(* IEC 61131-3 sources: STEPROBOT/docs/welder_r6_4/plc, 4 files *)

(* ---- GVL_WelderBridge.st ---- *)
{attribute 'qualified_only'}
VAR_GLOBAL PERSISTENT RETAIN
    // AC802 fixed MW registers require both persistence attributes.
    aCommand AT %MW7000 : ARRAY[0..31] OF WORD;
    wHeartbeat AT %MW7064 : WORD;
    aStatus AT %MW7200 : ARRAY[0..63] OF WORD;
END_VAR

VAR_GLOBAL
    // Local commissioning inputs; never write these over the PC command channel.
    xMappingConfirmed : BOOL := FALSE;
    xWeldPermit : BOOL := FALSE;
    // Drive from the real EtherCAT slave OP / working-counter-valid signal.
    // A constant TRUE is not a valid connection-health signal.
    xPdoOperational : BOOL := FALSE;
END_VAR

(* ---- GVL_Welders.st ---- *)
(* Reused legacy EtherCAT PDO variables. No fixed addresses or retained process outputs.
   Old Dxxx comments describe the source only; PC uses HR7000 / HR7200. *)
VAR_GLOBAL
    (* EtherCAT输出 → 焊机输入数据区 (32字节) *)
    g_byWeldOut : ARRAY[0..31] OF BYTE;
    (* EtherCAT输入 ← 焊机输出数据区 (32字节) *)
    g_byWeldIn : ARRAY[0..31] OF BYTE;

    (*
     * EtherCAT 映射别名。
     * InoProShop 的 I/O 映射器要求变量是单一标识符，不接受数组下标；
     * CommPoll 在这些别名与协议数组之间逐周期同步，协议字节编号保持不变。
     *)
    g_byWeldOutMap01 : BYTE;
    g_byWeldOutMap02 : BYTE;
    g_byWeldOutMap03 : BYTE;
    g_byWeldOutMap04 : BYTE;
    g_byWeldOutMap05 : BYTE;
    g_byWeldOutMap06 : BYTE;
    g_byWeldOutMap07 : BYTE;
    g_byWeldOutMap08 : BYTE;
    g_byWeldOutMap09 : BYTE;
    g_byWeldOutMap10 : BYTE;
    g_byWeldOutMap11 : BYTE;
    g_byWeldOutMap12 : BYTE;
    g_byWeldOutMap13 : BYTE;
    g_byWeldOutMap14 : BYTE;
    g_byWeldOutMap15 : BYTE;
    g_byWeldOutMap16 : BYTE;
    g_byWeldOutMap17 : BYTE;
    g_byWeldOutMap18 : BYTE;
    g_byWeldOutMap19 : BYTE;
    g_byWeldOutMap20 : BYTE;
    g_byWeldOutMap21 : BYTE;
    g_byWeldOutMap22 : BYTE;
    g_byWeldOutMap23 : BYTE;
    g_byWeldOutMap24 : BYTE;
    g_byWeldOutMap25 : BYTE;
    g_byWeldOutMap26 : BYTE;
    g_byWeldOutMap27 : BYTE;
    g_byWeldOutMap28 : BYTE;
    g_byWeldOutMap29 : BYTE;
    g_byWeldOutMap30 : BYTE;
    g_byWeldOutMap31 : BYTE;
    g_byWeldOutMap32 : BYTE;

    g_byWeldInMap01 : BYTE;
    g_byWeldInMap02 : BYTE;
    g_byWeldInMap03 : BYTE;
    g_byWeldInMap04 : BYTE;
    g_byWeldInMap05 : BYTE;
    g_byWeldInMap06 : BYTE;
    g_byWeldInMap07 : BYTE;
    g_byWeldInMap08 : BYTE;
    g_byWeldInMap09 : BYTE;
    g_byWeldInMap10 : BYTE;
    g_byWeldInMap11 : BYTE;
    g_byWeldInMap12 : BYTE;
    g_byWeldInMap13 : BYTE;
    g_byWeldInMap14 : BYTE;
    g_byWeldInMap15 : BYTE;
    g_byWeldInMap16 : BYTE;
    g_byWeldInMap17 : BYTE;
    g_byWeldInMap18 : BYTE;
    g_byWeldInMap19 : BYTE;
    g_byWeldInMap20 : BYTE;
    g_byWeldInMap21 : BYTE;
    g_byWeldInMap22 : BYTE;
    g_byWeldInMap23 : BYTE;
    g_byWeldInMap24 : BYTE;
    g_byWeldInMap25 : BYTE;
    g_byWeldInMap26 : BYTE;
    g_byWeldInMap27 : BYTE;
    g_byWeldInMap28 : BYTE;
    g_byWeldInMap29 : BYTE;
    g_byWeldInMap30 : BYTE;
    g_byWeldInMap31 : BYTE;
    g_byWeldInMap32 : BYTE;

	(* D520 | 激光距离 (原始INT值, 从%IW50读取) *)
	(* --- 激光距离原始值 --- *)
	g_iLaserDistanceRaw : INT;
END_VAR

VAR_GLOBAL

(* D300 | 控制标志位打包字 (PC通过Modbus读写, CommPoll每周期双向映射) *)
g_wWeldCtrlWord : UINT := 0;

(* D300 bit0 | 独立BOOL | 开始焊接 1=起弧 0=停弧 [危险, 高有效] *)
g_wWeldOn : BOOL := FALSE;

(* D300 bit1 | 独立BOOL | 机器人准备好, 高有效 *)
g_wRobotReady : BOOL := FALSE;
(* D300 bit2 | 独立BOOL | 检气, 高有效 *)
g_wGasCheck : BOOL := FALSE;

(* D300 bit3 | 独立BOOL | 热丝电源使能 1=ON 0=OFF *)
g_bHotWireEnable : BOOL := FALSE;

(* D300 bit4 | 独立BOOL | 热丝工作模式 0=DC 1=AC *)
g_bHotWireACMode : BOOL := FALSE;

(* D300 bit7 | 独立BOOL | 高频有无 0=高频 1=提升 *)
g_bHighFreqDisable : BOOL := FALSE;

(* D300 bit8 | 独立BOOL | 焊枪模式 0=水冷 1=气冷 *)
g_bGunCoolMode : BOOL := FALSE;

(* D302 | 协议Byte0 bit3-4 | 焊机操作模式 0=两步 1=四步 2=反复 *)
g_wWeldOperMode : UINT := 0;

(* D304 | 协议Byte0 bit5-7 | 焊机工作模式 0=直流恒流 1=直流脉冲 2=交流恒流 *)
(*                           3=交流脉冲 4=直流手弧焊 *)
g_wWeldWorkMode : UINT := 1;

(* D306 | 协议Byte11 | 通讯异常标志, 控制器填充, 默认0 *)
g_wCommErrorFlag : BYTE;

(* D414 | 协议Byte2 bit0-7 | 热丝频率, 范围20~100, 对应20~100Hz (直通) *)
g_wHotWireFreq : UINT := 50;

(* D416 | 协议Byte3 bit0-7 | 热丝电流给定, 范围0~200, 对应0~200A (直通) *)
g_wHotWireCurrent : UINT := 150;

(* D400 | 协议Byte4-5 | 给定电流, 实际A, 例: 100.0表示100.0A *)
(* CommPoll内部 ×10 → 协议值(范围40~4000, 对应4.0~400.0A), 占D400-D401 *)
g_wWeldCurrent : REAL := 100.0;

(* Local wire-feed axis parameters. Speeds are mm/s; delays are seconds.
   D412 and D1202 set the same automatic speed; a changed D1202 has priority.
   D410 > 0 overrides D2104 for axis 4 jog; zero uses D2104 for compatibility. *)
g_rWireStartDelay : REAL := 0.0;
g_rWireStopDelay : REAL := 0.0;
g_rWireJogSpeed : REAL := 0.0;
g_rWireAutoSpeed : REAL := 0.0;

(* D420 | 协议Byte13-14 | 前气时间, 实际s, 例: 5.0表示5.00s *)
(* CommPoll内部 ×100 → 协议值(范围1~999, 对应0.01~9.99s), 占D420-D421 *)
g_wFrontGasTime : REAL := 0.01;

(* D422 | 协议Byte15-16 | 延气时间, 实际s, 例: 3.0表示3.0s *)
(* CommPoll内部 ×10 → 协议值(范围1~600, 对应0.1~60.0s), 占D422-D423 *)
g_wTailGasTime : REAL := 0.2;

(* D424 | 协议Byte17 bit0-7 | 爬升时间, 实际s, 例: 5.0表示5.0s *)
(* CommPoll内部 ×10 → 协议值(范围1~100, 对应0.1~10.0s), 占D424-D425 *)
g_wRampUpTime : REAL := 0.5;

(* D426 | 协议Byte18 bit0-7 | 衰减时间, 实际s, 例: 5.0表示5.0s *)
(* CommPoll内部 ×10 → 协议值(范围1~150, 对应0.1~15.0s) *)
g_wRampDownTime : REAL := 0.2;

(* D428 | 协议Byte19 bit0-7 | 脉冲频率, 实际Hz, 例: 5.0表示5.0Hz *)
(* CommPoll内部 ×10 → 协议值(范围2~200, 对应0.2~20.0Hz), 占D428-D429 *)
g_wPulseFreq : REAL := 0.5;

(* D430 | 协议Byte20+22 bit4-7 | 占空比, 实际百分比, 例: 50.0表示50.0% *)
(* CommPoll内部 ×10 → 协议值(范围1~999, 对应0.1%~99.9%), 占D430-D431 *)
g_wDutyCycle : REAL := 50.0;

(* D432 | 协议Byte21+22 bit0-3 | 峰值电流, 实际A, 例: 150.0表示150.0A *)
(* CommPoll内部 ×10 → 协议值(范围50~4000, 对应5.0~400.0A), 占D432-D433 *)
g_wPeakCurrent : REAL := 100.0;

(* D434 | 协议Byte23-24 | 基值电流, 实际A, 例: 30.0表示30.0A *)
(* CommPoll内部 ×10 → 协议值(范围50~4000, 对应5.0~400.0A), 占D434-D435 *)
g_wBaseCurrent : REAL := 30.0;

(* D436 | 协议Byte25-26 | 起弧电流, 实际A, 例: 100.0表示100.0A *)
(* CommPoll内部 ×10 → 协议值(范围50~4000, 对应5.0~400.0A), 占D436-D437 *)
(* --- 协议 Byte 25-26: 起弧电流 (2字节小端, 低字节在前) --- *)
g_wArcStartCurrent : REAL := 5.0;

(* D438 | 协议Byte27-28 | 收弧电流, 实际A, 例: 100.0表示100.0A *)
(* CommPoll内部 ×10 → 协议值(范围50~4000, 对应5.0~400.0A), 占D438-D439 *)
(* --- 协议 Byte 27-28: 收弧电流 (2字节小端, 低字节在前) --- *)
g_wArcEndCurrent : REAL := 5.0;

(* D440 | 协议Byte29 bit0-7 | 交流频率, 范围40~250, 对应40~250Hz (直通) *)
(* --- 协议 Byte 29: 交流频率 --- *)
g_wACFreq : UINT := 40;

(* D442 | 协议Byte30 bit0-7 | 清理比例, 范围90~180, 对应40~-50 *)
(* 协议转换: Byte30 = -1 × D442 + 130 *)
(* 例: D442=90 → Byte30=40, D442=130 → Byte30=0, D442=180 → Byte30=-50 *)
(* --- 协议 Byte 30: 清理比例 --- *)
g_wCleanRatio : UINT := 90;

(* D444 | 协议Byte31 bit0-7 | 交流偏置, 范围90~180, 对应40~-50 *)
(* 协议转换: Byte31 = -1 × D444 + 130 *)
(* 例: D444=90 → Byte31=40, D444=130 → Byte31=0, D444=180 → Byte31=-50 *)
(* --- 协议 Byte 31: 交流偏置 --- *)
g_wACBias : UINT := 90;

(* D308 | 输入状态打包字 (PC通过Modbus读取, CommPoll每周期从独立BOOL组装) *)
g_wWeldStatusWord : UINT;

(* D308 bit0 | 独立BOOL | 引弧成功, 高有效 *)
g_bWeldArcOK : BOOL;

(* D308 bit1 | 独立BOOL | 焊机准备好, 高有效 *)
g_bWeldReady : BOOL;

(* D308 bit2 | 独立BOOL | 电流有无, 高有效 *)
g_bWeldHasCurrent : BOOL;

(* D308 bit3 | 独立BOOL | 焊枪开关异常, 高有效 *)
g_bGunSwitchFault : BOOL;

(* D308 bit4 | 独立BOOL | 焊机热保护, 高有效 *)
g_bWeldThermalProtect : BOOL;

(* D308 bit5 | 独立BOOL | 缺水保护, 高有效 *)
g_bWaterProtect : BOOL;

(* D308 bit6 | 独立BOOL | 热丝电源热保护, 高有效 *)
g_bWirePSThermal : BOOL;

(* D308 bit7 | 独立BOOL | 热丝电源通讯保护, 高有效, 控制器填充 *)
g_bWirePSCommFault : BOOL;

(* D308 bit8 | 独立BOOL | 组合报警, 包含焊枪开关/热保护/缺水/热丝电源故障 *)
g_bWeldFault : BOOL;

(* D500 | 焊机输入状态字 (16位打包, 详见位域定义) *)
g_wWeldInStatus : UINT;

(* D502-D503 | 协议输入Byte4-5 | 实际焊接电压, 0.1V分辨率 *)
(* --- 协议输入 Byte 4-5: 实际焊接电压 (2字节小端, 0.1V分辨率) --- *)
(* 范围: 0~1000 → 0~100.0V *)
g_rWeldVoltageAct : REAL;

(* D506-D507 | 协议输入Byte6-7 | 实际焊接电流, 0.1A分辨率 *)
(* --- 协议输入 Byte 6-7: 实际焊接电流 (2字节小端, 0.1A分辨率) --- *)
(* 范围: 0~400 → 0~400A *)
g_rWeldCurrentAct : REAL;

(* D510-D511 | 协议输入Byte8-9 | 实际热丝焊接电流, 10A分辨率 *)
(* --- 协议输入 Byte 8-9: 实际热丝焊接电流 (2字节小端, 10A分辨率) --- *)
(* 范围: 0~20 → 0~200A *)
g_rHotWireCurrentAct : REAL;

(* D518 | 协议输入Byte1原始值 | 报警码, 报警时记录协议输入Byte1原始值 *)
(* --- 报警原始字节 --- *)
g_rWeldFaultCode : UINT;

(* D522 | 激光距离 (实际距离mm, 原始值/100+50) *)
(* --- 激光距离实际值 --- *)
g_rLaserDistance : REAL := 50.0;

(* ================================================================= *)
(* 协议输入预留字节 (协议保留, 当前未使用)                               *)
(*   协议输入 Byte 2-3: 预留                                          *)
(*   协议输入 Byte 12:  预留                                          *)
(* ================================================================= *)

END_VAR

(* ---- PRG_WelderBridge.st ---- *)
PROGRAM PRG_WelderBridge
VAR
    aFrame : ARRAY[0..31] OF WORD;
    aParam : ARRAY[0..19] OF WORD;
    uiI : UINT;
    wCheck : WORD;
    uiScan : UINT;
    wPreviousHeartbeat : WORD;
    xHeartbeatSeen : BOOL;
    xHeartbeatEdge : BOOL;
    fbWatchdog : TON;
    xHostFresh : BOOL;
    xBasePermit : BOOL;
    xArcPermit : BOOL;
    xParametersValid : BOOL;
    xWasRunning : BOOL;
    xJobEnded : BOOL;
    udiOwner : UDINT;
    udiCurrentOwner : UDINT;
    udiRequest : UDINT;
    udiLastRequest : UDINT;
    udiRequestOwner : UDINT;
    udiRequestBoot : UDINT;
    udiBoot : UDINT;
    wResult : WORD;
    wError : WORD;
    wOperation : WORD;
    wControl : WORD;
    wApplied : WORD;
END_VAR

// Call once per scan, after PRG_RobotBridge. No other task writes the welder PDOs.
udiBoot := GVL_RobotBridgeRetain.udiBootCounter;
udiCurrentOwner := SHL(WORD_TO_UDINT(GVL_RobotBridge.aHostStatus[15]),16) OR WORD_TO_UDINT(GVL_RobotBridge.aHostStatus[16]);
IF udiCurrentOwner <> udiOwner THEN
    udiOwner := udiCurrentOwner; udiLastRequest := 0; wControl := 0;
    xHeartbeatSeen := FALSE; wPreviousHeartbeat := GVL_WelderBridge.wHeartbeat;
END_IF;
xHeartbeatEdge := GVL_WelderBridge.wHeartbeat <> wPreviousHeartbeat;
IF xHeartbeatEdge THEN
    wPreviousHeartbeat := GVL_WelderBridge.wHeartbeat; xHeartbeatSeen := TRUE;
END_IF;
fbWatchdog(IN := NOT xHeartbeatEdge, PT := T#1200ms);
xHostFresh := xHeartbeatSeen AND NOT fbWatchdog.Q AND GVL_RobotBridge.xHostRegistered AND GVL_RobotBridge.xHostAlive AND (udiOwner <> 0);
xBasePermit := xHostFresh AND GVL_WelderBridge.xMappingConfirmed AND GVL_WelderBridge.xWeldPermit AND GVL_WelderBridge.xPdoOperational
    AND GVL_RobotBridge.xRobotLinkOK AND GVL_RobotBridge.xRemotePermit
    AND NOT GVL_RobotBridge.xStopInterlock AND NOT GVL_RobotBridge.xRobotEmergency AND NOT GVL_RobotBridge.xRobotAlarm;
xArcPermit := xBasePermit AND GVL_RobotBridge.xRobotExternalAuto AND NOT GVL_RobotBridge.xRobotPaused;
xJobEnded := xWasRunning AND NOT GVL_RobotBridge.xRobotRunning;
xWasRunning := GVL_RobotBridge.xRobotRunning;
IF NOT xBasePermit THEN wControl := 0; END_IF;
IF NOT xArcPermit OR xJobEnded THEN wControl := wControl AND WORD#16#0006; END_IF;

// Snapshot the whole FC16 frame, then check checksum, identity and monotonic request.
FOR uiI := 0 TO 31 DO aFrame[uiI] := GVL_WelderBridge.aCommand[uiI]; END_FOR;
udiRequest := SHL(WORD_TO_UDINT(aFrame[2]),16) OR WORD_TO_UDINT(aFrame[3]);
udiRequestOwner := SHL(WORD_TO_UDINT(aFrame[4]),16) OR WORD_TO_UDINT(aFrame[5]);
udiRequestBoot := SHL(WORD_TO_UDINT(aFrame[6]),16) OR WORD_TO_UDINT(aFrame[7]);
wCheck := WORD#16#A55A;
FOR uiI := 0 TO 30 DO wCheck := wCheck XOR aFrame[uiI]; END_FOR;
IF (aFrame[0] = WORD#16#5742) AND (aFrame[1] = WORD#1) AND (wCheck = aFrame[31])
    AND (udiRequestOwner = udiOwner) AND (udiOwner <> 0) AND (udiRequestBoot = udiBoot)
    AND (udiRequest > udiLastRequest) THEN
    udiLastRequest := udiRequest; wOperation := aFrame[8]; wResult := 2; wError := 0;
    IF wOperation = WORD#3 THEN
        wControl := 0; wResult := 1;
    ELSIF NOT xBasePermit THEN
        wError := 1;
    ELSIF wOperation = WORD#1 THEN
        IF (aFrame[9] AND WORD#16#FFF0) <> 0 THEN wError := 2;
        ELSIF ((aFrame[9] AND WORD#16#0009) <> 0) AND NOT xArcPermit THEN wError := 3;
        ELSIF ((aFrame[9] AND WORD#16#0009) <> 0) AND (((aFrame[9] AND WORD#2) = 0) OR NOT GVL_Welders.g_bWeldReady OR GVL_Welders.g_bWeldFault) THEN wError := 4;
        ELSIF ((aFrame[9] AND WORD#1) <> 0) AND ((aFrame[9] AND WORD#4) <> 0) THEN wError := 5;
        ELSE wControl := aFrame[9]; wResult := 1;
        END_IF;
    ELSIF wOperation = WORD#2 THEN
        IF wControl <> 0 THEN wError := 6;
        ELSE
            FOR uiI := 0 TO 19 DO aParam[uiI] := aFrame[10+uiI]; END_FOR;
            xParametersValid := TRUE;
            IF (aParam[0] < WORD#0) OR (aParam[0] > WORD#2) THEN xParametersValid := FALSE; END_IF;
            IF (aParam[1] < WORD#0) OR (aParam[1] > WORD#4) THEN xParametersValid := FALSE; END_IF;
            IF (aParam[2] < WORD#40) OR (aParam[2] > WORD#4000) THEN xParametersValid := FALSE; END_IF;
            IF (aParam[3] < WORD#20) OR (aParam[3] > WORD#100) THEN xParametersValid := FALSE; END_IF;
            IF (aParam[4] < WORD#0) OR (aParam[4] > WORD#200) THEN xParametersValid := FALSE; END_IF;
            IF (aParam[5] < WORD#1) OR (aParam[5] > WORD#999) THEN xParametersValid := FALSE; END_IF;
            IF (aParam[6] < WORD#1) OR (aParam[6] > WORD#600) THEN xParametersValid := FALSE; END_IF;
            IF (aParam[7] < WORD#1) OR (aParam[7] > WORD#100) THEN xParametersValid := FALSE; END_IF;
            IF (aParam[8] < WORD#1) OR (aParam[8] > WORD#150) THEN xParametersValid := FALSE; END_IF;
            IF (aParam[9] < WORD#2) OR (aParam[9] > WORD#200) THEN xParametersValid := FALSE; END_IF;
            IF (aParam[10] < WORD#1) OR (aParam[10] > WORD#999) THEN xParametersValid := FALSE; END_IF;
            IF (aParam[11] < WORD#50) OR (aParam[11] > WORD#4000) THEN xParametersValid := FALSE; END_IF;
            IF (aParam[12] < WORD#50) OR (aParam[12] > WORD#4000) THEN xParametersValid := FALSE; END_IF;
            IF (aParam[13] < WORD#50) OR (aParam[13] > WORD#4000) THEN xParametersValid := FALSE; END_IF;
            IF (aParam[14] < WORD#50) OR (aParam[14] > WORD#4000) THEN xParametersValid := FALSE; END_IF;
            IF (aParam[15] < WORD#40) OR (aParam[15] > WORD#250) THEN xParametersValid := FALSE; END_IF;
            IF (aParam[16] < WORD#90) OR (aParam[16] > WORD#180) THEN xParametersValid := FALSE; END_IF;
            IF (aParam[17] < WORD#90) OR (aParam[17] > WORD#180) THEN xParametersValid := FALSE; END_IF;
            IF (aParam[18] > WORD#7) OR (aParam[19] <> 0) THEN xParametersValid := FALSE; END_IF;
            IF NOT xParametersValid THEN wError := 7;
            ELSE
                GVL_Welders.g_wWeldOperMode := WORD_TO_UINT(aParam[0]);
                GVL_Welders.g_wWeldWorkMode := WORD_TO_UINT(aParam[1]);
                GVL_Welders.g_wWeldCurrent := UINT_TO_REAL(WORD_TO_UINT(aParam[2])) / 10.0;
                GVL_Welders.g_wHotWireFreq := WORD_TO_UINT(aParam[3]);
                GVL_Welders.g_wHotWireCurrent := WORD_TO_UINT(aParam[4]);
                GVL_Welders.g_wFrontGasTime := UINT_TO_REAL(WORD_TO_UINT(aParam[5])) / 100.0;
                GVL_Welders.g_wTailGasTime := UINT_TO_REAL(WORD_TO_UINT(aParam[6])) / 10.0;
                GVL_Welders.g_wRampUpTime := UINT_TO_REAL(WORD_TO_UINT(aParam[7])) / 10.0;
                GVL_Welders.g_wRampDownTime := UINT_TO_REAL(WORD_TO_UINT(aParam[8])) / 10.0;
                GVL_Welders.g_wPulseFreq := UINT_TO_REAL(WORD_TO_UINT(aParam[9])) / 10.0;
                GVL_Welders.g_wDutyCycle := UINT_TO_REAL(WORD_TO_UINT(aParam[10])) / 10.0;
                GVL_Welders.g_wPeakCurrent := UINT_TO_REAL(WORD_TO_UINT(aParam[11])) / 10.0;
                GVL_Welders.g_wBaseCurrent := UINT_TO_REAL(WORD_TO_UINT(aParam[12])) / 10.0;
                GVL_Welders.g_wArcStartCurrent := UINT_TO_REAL(WORD_TO_UINT(aParam[13])) / 10.0;
                GVL_Welders.g_wArcEndCurrent := UINT_TO_REAL(WORD_TO_UINT(aParam[14])) / 10.0;
                GVL_Welders.g_wACFreq := WORD_TO_UINT(aParam[15]);
                GVL_Welders.g_wCleanRatio := WORD_TO_UINT(aParam[16]);
                GVL_Welders.g_wACBias := WORD_TO_UINT(aParam[17]);
                GVL_Welders.g_bHotWireACMode := (aParam[18] AND WORD#1) <> 0;
                GVL_Welders.g_bHighFreqDisable := (aParam[18] AND WORD#2) <> 0;
                GVL_Welders.g_bGunCoolMode := (aParam[18] AND WORD#4) <> 0;
                wResult := 1;
            END_IF;
        END_IF;
    ELSE wError := 8;
    END_IF;
END_IF;
GVL_Welders.g_wWeldOn := (wControl AND WORD#1) <> 0;
GVL_Welders.g_wRobotReady := (wControl AND WORD#2) <> 0;
GVL_Welders.g_wGasCheck := (wControl AND WORD#4) <> 0;
GVL_Welders.g_bHotWireEnable := (wControl AND WORD#8) <> 0;
PRG_WelderIo();
// Same-scan PDO input interlock; never restore an arc after a fault clears.
IF NOT GVL_Welders.g_bWeldReady OR GVL_Welders.g_bWeldFault THEN
    wControl := wControl AND WORD#16#0006;
    GVL_Welders.g_wWeldOn := FALSE; GVL_Welders.g_bHotWireEnable := FALSE;
    GVL_Welders.g_byWeldOutMap01 := GVL_Welders.g_byWeldOutMap01 AND BYTE#16#FE;
    GVL_Welders.g_byWeldOutMap02 := GVL_Welders.g_byWeldOutMap02 AND BYTE#16#FE;
END_IF;
wApplied := wControl;
GVL_Welders.g_wWeldCtrlWord := WORD_TO_UINT(wApplied);
uiScan := uiScan + UINT#1;
GVL_WelderBridge.aStatus[0] := WORD#16#5742;
GVL_WelderBridge.aStatus[1] := 1;
GVL_WelderBridge.aStatus[2] := UINT_TO_WORD(uiScan);
GVL_WelderBridge.aStatus[3] := 1;
IF GVL_WelderBridge.xMappingConfirmed THEN GVL_WelderBridge.aStatus[3] := GVL_WelderBridge.aStatus[3] OR WORD#2; END_IF;
IF GVL_WelderBridge.xPdoOperational THEN GVL_WelderBridge.aStatus[3] := GVL_WelderBridge.aStatus[3] OR WORD#4; END_IF;
IF xBasePermit THEN GVL_WelderBridge.aStatus[3] := GVL_WelderBridge.aStatus[3] OR WORD#8; END_IF;
IF xHostFresh THEN GVL_WelderBridge.aStatus[3] := GVL_WelderBridge.aStatus[3] OR WORD#16; END_IF;
IF xArcPermit THEN GVL_WelderBridge.aStatus[3] := GVL_WelderBridge.aStatus[3] OR WORD#32; END_IF;
GVL_WelderBridge.aStatus[4] := UDINT_TO_WORD(SHR(udiBoot,16));
GVL_WelderBridge.aStatus[5] := UDINT_TO_WORD(udiBoot AND UDINT#65535);
GVL_WelderBridge.aStatus[6] := UDINT_TO_WORD(SHR(udiLastRequest,16));
GVL_WelderBridge.aStatus[7] := UDINT_TO_WORD(udiLastRequest AND UDINT#65535);
GVL_WelderBridge.aStatus[8] := wResult;
GVL_WelderBridge.aStatus[9] := wError;
GVL_WelderBridge.aStatus[10] := wApplied;
GVL_WelderBridge.aStatus[11] := UINT_TO_WORD(GVL_Welders.g_wWeldInStatus);
GVL_WelderBridge.aStatus[12] := UINT_TO_WORD(GVL_Welders.g_rWeldFaultCode);
GVL_WelderBridge.aStatus[13] := wOperation;
GVL_WelderBridge.aStatus[14] := UDINT_TO_WORD(SHR(udiOwner,16));
GVL_WelderBridge.aStatus[15] := UDINT_TO_WORD(udiOwner AND UDINT#65535);
GVL_WelderBridge.aStatus[16] := REAL_TO_WORD(LIMIT(0.0,GVL_Welders.g_rWeldVoltageAct*10.0,65535.0));
GVL_WelderBridge.aStatus[17] := REAL_TO_WORD(LIMIT(0.0,GVL_Welders.g_rWeldCurrentAct*10.0,65535.0));
GVL_WelderBridge.aStatus[18] := REAL_TO_WORD(LIMIT(0.0,GVL_Welders.g_rHotWireCurrentAct*10.0,65535.0));
GVL_WelderBridge.aStatus[19] := GVL_WelderBridge.wHeartbeat;
GVL_WelderBridge.aStatus[20] := UINT_TO_WORD(GVL_Welders.g_wWeldOperMode);
GVL_WelderBridge.aStatus[21] := UINT_TO_WORD(GVL_Welders.g_wWeldWorkMode);
GVL_WelderBridge.aStatus[22] := REAL_TO_WORD(GVL_Welders.g_wWeldCurrent * 10.0);
GVL_WelderBridge.aStatus[23] := UINT_TO_WORD(GVL_Welders.g_wHotWireFreq);
GVL_WelderBridge.aStatus[24] := UINT_TO_WORD(GVL_Welders.g_wHotWireCurrent);
GVL_WelderBridge.aStatus[25] := REAL_TO_WORD(GVL_Welders.g_wFrontGasTime * 100.0);
GVL_WelderBridge.aStatus[26] := REAL_TO_WORD(GVL_Welders.g_wTailGasTime * 10.0);
GVL_WelderBridge.aStatus[27] := REAL_TO_WORD(GVL_Welders.g_wRampUpTime * 10.0);
GVL_WelderBridge.aStatus[28] := REAL_TO_WORD(GVL_Welders.g_wRampDownTime * 10.0);
GVL_WelderBridge.aStatus[29] := REAL_TO_WORD(GVL_Welders.g_wPulseFreq * 10.0);
GVL_WelderBridge.aStatus[30] := REAL_TO_WORD(GVL_Welders.g_wDutyCycle * 10.0);
GVL_WelderBridge.aStatus[31] := REAL_TO_WORD(GVL_Welders.g_wPeakCurrent * 10.0);
GVL_WelderBridge.aStatus[32] := REAL_TO_WORD(GVL_Welders.g_wBaseCurrent * 10.0);
GVL_WelderBridge.aStatus[33] := REAL_TO_WORD(GVL_Welders.g_wArcStartCurrent * 10.0);
GVL_WelderBridge.aStatus[34] := REAL_TO_WORD(GVL_Welders.g_wArcEndCurrent * 10.0);
GVL_WelderBridge.aStatus[35] := UINT_TO_WORD(GVL_Welders.g_wACFreq);
GVL_WelderBridge.aStatus[36] := UINT_TO_WORD(GVL_Welders.g_wCleanRatio);
GVL_WelderBridge.aStatus[37] := UINT_TO_WORD(GVL_Welders.g_wACBias);
IF GVL_WelderBridge.xWeldPermit THEN GVL_WelderBridge.aStatus[3] := GVL_WelderBridge.aStatus[3] OR WORD#64; END_IF;
GVL_WelderBridge.aStatus[38] := 0;
IF GVL_Welders.g_bHotWireACMode THEN GVL_WelderBridge.aStatus[38] := GVL_WelderBridge.aStatus[38] OR WORD#1; END_IF;
IF GVL_Welders.g_bHighFreqDisable THEN GVL_WelderBridge.aStatus[38] := GVL_WelderBridge.aStatus[38] OR WORD#2; END_IF;
IF GVL_Welders.g_bGunCoolMode THEN GVL_WelderBridge.aStatus[38] := GVL_WelderBridge.aStatus[38] OR WORD#4; END_IF;
GVL_WelderBridge.aStatus[39] := 0;
FOR uiI := 0 TO 15 DO
    GVL_WelderBridge.aStatus[40+uiI] := BYTE_TO_WORD(GVL_Welders.g_byWeldIn[uiI*2]) OR SHL(BYTE_TO_WORD(GVL_Welders.g_byWeldIn[uiI*2+1]),8);
END_FOR;
FOR uiI := 56 TO 63 DO GVL_WelderBridge.aStatus[uiI] := 0; END_FOR;
END_PROGRAM

(* ---- PRG_WelderIo.st ---- *)
(* Reused from lower.project CommPoll: unchanged PDO byte encoding and feedback units. *)
PROGRAM PRG_WelderIo
VAR
    nTempU16 : UINT;
    nTempI16 : INT;
    byTemp : BYTE;
END_VAR
(* ================================================================ *)
(* 焊机输出 (协议: 焊机的输入数据区, PLC写→焊机读)                    *)
(* GVL_Welders.g_byWeldOut[0..31] → EtherCAT输出 → 焊机                        *)
(* ================================================================ *)

(* ===== 协议 Byte 0: 控制位 ===== *)
(* bit0(1):  开始焊接 1=起弧 0=停弧                                  *)
(* bit1(2):  机器人准备好 高有效                                      *)
(* bit2(3):  检气 高有效                                              *)
(* bit3-4:   焊机操作模式 00=两步 01=四步 10=反复                     *)
(* bit5-7:   焊机工作模式 000=直流恒流 001=直流脉冲 010=交流恒流       *)
(*           011=交流脉冲 100=直流手弧焊                               *)
byTemp := 0;
IF GVL_Welders.g_wWeldOn THEN byTemp := byTemp OR 16#01; END_IF;
IF GVL_Welders.g_wRobotReady THEN byTemp := byTemp OR 16#02; END_IF;
IF GVL_Welders.g_wGasCheck THEN byTemp := byTemp OR 16#04; END_IF;
nTempU16 := LIMIT(UINT#0, GVL_Welders.g_wWeldOperMode, UINT#2);
byTemp := byTemp OR SHL(UINT_TO_BYTE(nTempU16), 3);
nTempU16 := LIMIT(UINT#0, GVL_Welders.g_wWeldWorkMode, UINT#4);
byTemp := byTemp OR SHL(UINT_TO_BYTE(nTempU16), 5);
GVL_Welders.g_byWeldOut[0] := byTemp;

(* ===== 协议 Byte 1: 辅助控制位 ===== *)
(* bit0(9):  热丝电源使能 1=ON 0=OFF                                  *)
(* bit1(10): 热丝工作模式 0=DC 1=AC                                   *)
(* bit2(11): 备用                                                     *)
(* bit3(12): 点动送丝 (已移除, 送丝通过轴控制) *)
(* bit4(13): 点动抽丝 (已移除, 送丝通过轴控制) *)
(* bit5(14): 备用                                                     *)
(* bit6(15): 高频有无 0=高频 1=提升                                   *)
(* bit7(16): 焊枪模式 0=水冷 1=气冷                                   *)
byTemp := 0;
IF GVL_Welders.g_bHotWireEnable THEN byTemp := byTemp OR 16#01; END_IF;
IF GVL_Welders.g_bHotWireACMode THEN byTemp := byTemp OR 16#02; END_IF;
IF GVL_Welders.g_bHighFreqDisable THEN byTemp := byTemp OR 16#40; END_IF;
IF GVL_Welders.g_bGunCoolMode THEN byTemp := byTemp OR 16#80; END_IF;
GVL_Welders.g_byWeldOut[1] := byTemp;

(* ===== 协议 Byte 2: 热丝频率 ===== *)
(* 范围: 20-100 对应20~100Hz (1字节) *)
GVL_Welders.g_byWeldOut[2] := UINT_TO_BYTE(LIMIT(UINT#20, GVL_Welders.g_wHotWireFreq, UINT#100));

(* ===== 协议 Byte 3: 热丝电流给定 ===== *)
(* 范围: 0-200 对应0~200A (1字节) *)
GVL_Welders.g_byWeldOut[3] := UINT_TO_BYTE(LIMIT(UINT#0, GVL_Welders.g_wHotWireCurrent, UINT#200));

(* ===== 协议 Byte 4-5: 给定电流 (2字节小端, 低字节在前) ===== *)
(* 范围: 40-4000 对应4.0~400.0A *)
nTempU16 := REAL_TO_UINT(LIMIT(4.0, GVL_Welders.g_wWeldCurrent, 400.0)*10.0);

GVL_Welders.g_byWeldOut[4] := UINT_TO_BYTE(UINT_TO_USINT(nTempU16 MOD 256));
GVL_Welders.g_byWeldOut[5] := UINT_TO_BYTE(UINT_TO_USINT(nTempU16 / 256));

(* ===== 协议 Byte 6: 送丝速度 (已移除, 送丝通过轴控制, 写0) ===== *)
GVL_Welders.g_byWeldOut[6] := 0;

(* ===== 协议 Byte 7: 起弧延迟送丝时间 (已移除, 写0) ===== *)
GVL_Welders.g_byWeldOut[7] := 0;

(* ===== 协议 Byte 8: 熄弧滞后送丝时间 (已移除, 写0) ===== *)
GVL_Welders.g_byWeldOut[8] := 0;

(* ===== 协议 Byte 9: 熄弧回抽丝长度 (已移除, 写0) ===== *)
GVL_Welders.g_byWeldOut[9] := 0;

(* ===== 协议 Byte 10: 点动送丝速度 (已移除, 送丝通过轴控制, 写0) ===== *)
GVL_Welders.g_byWeldOut[10] := 0;

(* ===== 协议 Byte 11: 通讯异常标志 (控制器填充) ===== *)
GVL_Welders.g_byWeldOut[11] := GVL_Welders.g_wCommErrorFlag;

(* ===== 协议 Byte 12: 慢送丝速度 (已移除, 送丝通过轴控制, 写0) ===== *)
GVL_Welders.g_byWeldOut[12] := 0;

(* ===== 协议 Byte 13-14: 前气时间 (2字节小端, 低字节在前) ===== *)
(* 范围: 1-999 对应0.01~9.99s *)
nTempU16 := REAL_TO_UINT(LIMIT(0.01, GVL_Welders.g_wFrontGasTime, 9.99)*100.0);
GVL_Welders.g_byWeldOut[13] := UINT_TO_BYTE(UINT_TO_USINT(nTempU16 MOD 256));
GVL_Welders.g_byWeldOut[14] := UINT_TO_BYTE(UINT_TO_USINT(nTempU16 / 256));

(* ===== 协议 Byte 15-16: 延气时间 (2字节小端, 低字节在前) ===== *)
(* 范围: 1-600 对应0.1~60.0s *)
nTempU16 := REAL_TO_UINT(LIMIT(0.1, GVL_Welders.g_wTailGasTime, 60.0)*10.0);
GVL_Welders.g_byWeldOut[15] := UINT_TO_BYTE(UINT_TO_USINT(nTempU16 MOD 256));
GVL_Welders.g_byWeldOut[16] := UINT_TO_BYTE(UINT_TO_USINT(nTempU16 / 256));

(* ===== 协议 Byte 17: 爬升时间 ===== *)
(* 范围: 1-100 对应0.1~10.0s (1字节) *)
GVL_Welders.g_byWeldOut[17] := UINT_TO_BYTE(REAL_TO_UINT(LIMIT(0.1, GVL_Welders.g_wRampUpTime, 10.0)*10.0));

(* ===== 协议 Byte 18: 衰减时间 ===== *)
(* 范围: 1-150 对应0.1~15.0s (1字节) *)
GVL_Welders.g_byWeldOut[18] := UINT_TO_BYTE(REAL_TO_UINT(LIMIT(0.1, GVL_Welders.g_wRampDownTime, 15.0)*10.0));

(* ===== 协议 Byte 19: 脉冲频率 ===== *)
(* 范围: 2-200 对应0.2~20.0Hz (1字节) *)
GVL_Welders.g_byWeldOut[19] := UINT_TO_BYTE(REAL_TO_UINT(LIMIT(0.2, GVL_Welders.g_wPulseFreq, 20.0)*10.0));

(* ===== 协议 Byte 20-22: 占空比 + 峰值电流 (交叉编排) ===== *)
(* 占空比: Byte20=低字节, Byte22 bit4-7=高字节低4位 (范围1-999, 12位) *)
(* 峰值电流: Byte21=低字节, Byte22 bit0-3=高字节低4位 (范围50-4000, 12位) *)
(* 占空比 = [Byte22 bit7:4][Byte20] *)
(* 峰值电流 = [Byte22 bit3:0][Byte21] *)
nTempU16 := REAL_TO_UINT(LIMIT(0.1, GVL_Welders.g_wDutyCycle, 99.9)*10.0);
GVL_Welders.g_byWeldOut[20] := UINT_TO_BYTE(UINT_TO_USINT(nTempU16 MOD 256));
GVL_Welders.g_byWeldOut[21] := UINT_TO_BYTE(UINT_TO_USINT(REAL_TO_UINT(LIMIT(5.0, GVL_Welders.g_wPeakCurrent, 400.0)*10.0) MOD 256));
byTemp := 0;
byTemp := byTemp OR SHL(UINT_TO_BYTE(UINT_TO_USINT(nTempU16 / 256)) AND 16#0F, 4);
byTemp := byTemp OR (UINT_TO_BYTE(UINT_TO_USINT(REAL_TO_UINT(LIMIT(5.0, GVL_Welders.g_wPeakCurrent, 400.0)*10.0) / 256)) AND 16#0F);
GVL_Welders.g_byWeldOut[22] := byTemp;

(* ===== 协议 Byte 23-24: 基值电流 (2字节小端, 低字节在前) ===== *)
(* 范围: 50-4000 对应5.0~400.0A *)
nTempU16 := REAL_TO_UINT(LIMIT(5.0, GVL_Welders.g_wBaseCurrent, 400.0)*10.0);
GVL_Welders.g_byWeldOut[23] := UINT_TO_BYTE(UINT_TO_USINT(nTempU16 MOD 256));
GVL_Welders.g_byWeldOut[24] := UINT_TO_BYTE(UINT_TO_USINT(nTempU16 / 256));

(* ===== 协议 Byte 25-26: 起弧电流 (2字节小端, 低字节在前) ===== *)
(* 范围: 50-4000 对应5.0~400.0A *)
nTempU16 := REAL_TO_UINT(LIMIT(5.0, GVL_Welders.g_wArcStartCurrent, 400.0)*10.0);
GVL_Welders.g_byWeldOut[25] := UINT_TO_BYTE(UINT_TO_USINT(nTempU16 MOD 256));
GVL_Welders.g_byWeldOut[26] := UINT_TO_BYTE(UINT_TO_USINT(nTempU16 / 256));

(* ===== 协议 Byte 27-28: 收弧电流 (2字节小端, 低字节在前) ===== *)
(* 范围: 50-4000 对应5.0~400.0A *)
nTempU16 := REAL_TO_UINT(LIMIT(5.0, GVL_Welders.g_wArcEndCurrent, 400.0)*10.0);
GVL_Welders.g_byWeldOut[27] := UINT_TO_BYTE(UINT_TO_USINT(nTempU16 MOD 256));
GVL_Welders.g_byWeldOut[28] := UINT_TO_BYTE(UINT_TO_USINT(nTempU16 / 256));

(* ===== 协议 Byte 29: 交流频率 ===== *)
(* 范围: 40-250 对应40-250Hz (1字节) *)
GVL_Welders.g_byWeldOut[29] := UINT_TO_BYTE(LIMIT(UINT#40, GVL_Welders.g_wACFreq, UINT#250));

(* ===== 协议 Byte 30: 清理比例 ===== *)
(* 范围: 90-180 对应40~-50 (1字节) *)
nTempI16 := 130 - UINT_TO_INT(LIMIT(UINT#90, GVL_Welders.g_wCleanRatio, UINT#180));
GVL_Welders.g_byWeldOut[30] := INT_TO_BYTE(nTempI16);

(* ===== 协议 Byte 31: 交流偏置 ===== *)
(* 范围: 90-180 对应40~-50 (1字节) *)
nTempI16 := 130 - UINT_TO_INT(LIMIT(UINT#90, GVL_Welders.g_wACBias, UINT#180));
GVL_Welders.g_byWeldOut[31] := INT_TO_BYTE(nTempI16);

(* ================================================================ *)
(* 焊机输入 (协议: 焊机输出数据区, 焊机写→PLC读)                      *)
(* GVL_Welders.g_byWeldIn[0..31] ← EtherCAT输入 ← 焊机                          *)
(* ================================================================ *)

(* ===== 协议输入 Byte 0: 状态位 ===== *)
(* bit0: 引弧成功 高有效                                              *)
(* bit1: 焊机准备好 高有效                                            *)
(* bit2: 预留                                                         *)
(* bit3: 电流有无 高有效                                              *)
(* EtherCAT 输入映射别名 → 协议数组。保持原有 Byte 0..31 定义。 *)
GVL_Welders.g_byWeldIn[0] := GVL_Welders.g_byWeldInMap01;
GVL_Welders.g_byWeldIn[1] := GVL_Welders.g_byWeldInMap02;
GVL_Welders.g_byWeldIn[2] := GVL_Welders.g_byWeldInMap03;
GVL_Welders.g_byWeldIn[3] := GVL_Welders.g_byWeldInMap04;
GVL_Welders.g_byWeldIn[4] := GVL_Welders.g_byWeldInMap05;
GVL_Welders.g_byWeldIn[5] := GVL_Welders.g_byWeldInMap06;
GVL_Welders.g_byWeldIn[6] := GVL_Welders.g_byWeldInMap07;
GVL_Welders.g_byWeldIn[7] := GVL_Welders.g_byWeldInMap08;
GVL_Welders.g_byWeldIn[8] := GVL_Welders.g_byWeldInMap09;
GVL_Welders.g_byWeldIn[9] := GVL_Welders.g_byWeldInMap10;
GVL_Welders.g_byWeldIn[10] := GVL_Welders.g_byWeldInMap11;
GVL_Welders.g_byWeldIn[11] := GVL_Welders.g_byWeldInMap12;
GVL_Welders.g_byWeldIn[12] := GVL_Welders.g_byWeldInMap13;
GVL_Welders.g_byWeldIn[13] := GVL_Welders.g_byWeldInMap14;
GVL_Welders.g_byWeldIn[14] := GVL_Welders.g_byWeldInMap15;
GVL_Welders.g_byWeldIn[15] := GVL_Welders.g_byWeldInMap16;
GVL_Welders.g_byWeldIn[16] := GVL_Welders.g_byWeldInMap17;
GVL_Welders.g_byWeldIn[17] := GVL_Welders.g_byWeldInMap18;
GVL_Welders.g_byWeldIn[18] := GVL_Welders.g_byWeldInMap19;
GVL_Welders.g_byWeldIn[19] := GVL_Welders.g_byWeldInMap20;
GVL_Welders.g_byWeldIn[20] := GVL_Welders.g_byWeldInMap21;
GVL_Welders.g_byWeldIn[21] := GVL_Welders.g_byWeldInMap22;
GVL_Welders.g_byWeldIn[22] := GVL_Welders.g_byWeldInMap23;
GVL_Welders.g_byWeldIn[23] := GVL_Welders.g_byWeldInMap24;
GVL_Welders.g_byWeldIn[24] := GVL_Welders.g_byWeldInMap25;
GVL_Welders.g_byWeldIn[25] := GVL_Welders.g_byWeldInMap26;
GVL_Welders.g_byWeldIn[26] := GVL_Welders.g_byWeldInMap27;
GVL_Welders.g_byWeldIn[27] := GVL_Welders.g_byWeldInMap28;
GVL_Welders.g_byWeldIn[28] := GVL_Welders.g_byWeldInMap29;
GVL_Welders.g_byWeldIn[29] := GVL_Welders.g_byWeldInMap30;
GVL_Welders.g_byWeldIn[30] := GVL_Welders.g_byWeldInMap31;
GVL_Welders.g_byWeldIn[31] := GVL_Welders.g_byWeldInMap32;

GVL_Welders.g_bWeldArcOK      := (GVL_Welders.g_byWeldIn[0] AND 16#01) <> 0;
GVL_Welders.g_bWeldReady      := (GVL_Welders.g_byWeldIn[0] AND 16#02) <> 0;
GVL_Welders.g_bWeldHasCurrent     := (GVL_Welders.g_byWeldIn[0] AND 16#08) <> 0;

(* ===== 协议输入 Byte 1: 报警位 ===== *)
(* bit0: 预留                                                         *)
(* bit1: 焊枪开关异常 高有效                                          *)
(* bit2: 焊机热保护 高有效                                            *)
(* bit3: 缺水保护 高有效                                              *)
(* bit4: 热丝电源热保护 高有效                                        *)
(* bit5: 热丝电源通讯保护 高有效 (控制器填充)                          *)
GVL_Welders.g_bGunSwitchFault    := (GVL_Welders.g_byWeldIn[1] AND 16#02) <> 0;
GVL_Welders.g_bWeldThermalProtect := (GVL_Welders.g_byWeldIn[1] AND 16#04) <> 0;
GVL_Welders.g_bWaterProtect   := (GVL_Welders.g_byWeldIn[1] AND 16#08) <> 0;
GVL_Welders.g_bWirePSThermal  := (GVL_Welders.g_byWeldIn[1] AND 16#10) <> 0;
GVL_Welders.g_bWirePSCommFault:= (GVL_Welders.g_byWeldIn[1] AND 16#20) <> 0;

(* ===== 报警组合 ===== *)
GVL_Welders.g_bWeldFault := GVL_Welders.g_bWeldThermalProtect
              OR GVL_Welders.g_bGunSwitchFault
              OR GVL_Welders.g_bWaterProtect
              OR GVL_Welders.g_bWirePSThermal
              OR GVL_Welders.g_bWirePSCommFault;

IF GVL_Welders.g_bWeldFault THEN
    GVL_Welders.g_rWeldFaultCode := BYTE_TO_UINT(GVL_Welders.g_byWeldIn[1]);
ELSE
    GVL_Welders.g_rWeldFaultCode := 0;
END_IF;

IF NOT GVL_Welders.g_bWeldReady OR GVL_Welders.g_bWeldFault THEN
    GVL_Welders.g_wWeldOn := FALSE;
    GVL_Welders.g_wWeldCtrlWord := GVL_Welders.g_wWeldCtrlWord AND 16#FFFE;
    GVL_Welders.g_byWeldOut[0] := GVL_Welders.g_byWeldOut[0] AND 16#FE;
END_IF;

(* ===== EtherCAT 输出映射别名同步 ===== *)
(* 放在未就绪/故障联锁之后，确保停弧命令在本周期立即写入PDO。 *)
GVL_Welders.g_byWeldOutMap01 := GVL_Welders.g_byWeldOut[0];
GVL_Welders.g_byWeldOutMap02 := GVL_Welders.g_byWeldOut[1];
GVL_Welders.g_byWeldOutMap03 := GVL_Welders.g_byWeldOut[2];
GVL_Welders.g_byWeldOutMap04 := GVL_Welders.g_byWeldOut[3];
GVL_Welders.g_byWeldOutMap05 := GVL_Welders.g_byWeldOut[4];
GVL_Welders.g_byWeldOutMap06 := GVL_Welders.g_byWeldOut[5];
GVL_Welders.g_byWeldOutMap07 := GVL_Welders.g_byWeldOut[6];
GVL_Welders.g_byWeldOutMap08 := GVL_Welders.g_byWeldOut[7];
GVL_Welders.g_byWeldOutMap09 := GVL_Welders.g_byWeldOut[8];
GVL_Welders.g_byWeldOutMap10 := GVL_Welders.g_byWeldOut[9];
GVL_Welders.g_byWeldOutMap11 := GVL_Welders.g_byWeldOut[10];
GVL_Welders.g_byWeldOutMap12 := GVL_Welders.g_byWeldOut[11];
GVL_Welders.g_byWeldOutMap13 := GVL_Welders.g_byWeldOut[12];
GVL_Welders.g_byWeldOutMap14 := GVL_Welders.g_byWeldOut[13];
GVL_Welders.g_byWeldOutMap15 := GVL_Welders.g_byWeldOut[14];
GVL_Welders.g_byWeldOutMap16 := GVL_Welders.g_byWeldOut[15];
GVL_Welders.g_byWeldOutMap17 := GVL_Welders.g_byWeldOut[16];
GVL_Welders.g_byWeldOutMap18 := GVL_Welders.g_byWeldOut[17];
GVL_Welders.g_byWeldOutMap19 := GVL_Welders.g_byWeldOut[18];
GVL_Welders.g_byWeldOutMap20 := GVL_Welders.g_byWeldOut[19];
GVL_Welders.g_byWeldOutMap21 := GVL_Welders.g_byWeldOut[20];
GVL_Welders.g_byWeldOutMap22 := GVL_Welders.g_byWeldOut[21];
GVL_Welders.g_byWeldOutMap23 := GVL_Welders.g_byWeldOut[22];
GVL_Welders.g_byWeldOutMap24 := GVL_Welders.g_byWeldOut[23];
GVL_Welders.g_byWeldOutMap25 := GVL_Welders.g_byWeldOut[24];
GVL_Welders.g_byWeldOutMap26 := GVL_Welders.g_byWeldOut[25];
GVL_Welders.g_byWeldOutMap27 := GVL_Welders.g_byWeldOut[26];
GVL_Welders.g_byWeldOutMap28 := GVL_Welders.g_byWeldOut[27];
GVL_Welders.g_byWeldOutMap29 := GVL_Welders.g_byWeldOut[28];
GVL_Welders.g_byWeldOutMap30 := GVL_Welders.g_byWeldOut[29];
GVL_Welders.g_byWeldOutMap31 := GVL_Welders.g_byWeldOut[30];
GVL_Welders.g_byWeldOutMap32 := GVL_Welders.g_byWeldOut[31];

(* ===== 协议输入 Byte 4-5: 实际焊接电压 (2字节小端, 0.1V分辨率) ===== *)
(* 范围: 0-1000 对应0~100.0V *)
nTempU16 := BYTE_TO_UINT(GVL_Welders.g_byWeldIn[4]) + BYTE_TO_UINT(GVL_Welders.g_byWeldIn[5]) * 256;
GVL_Welders.g_rWeldVoltageAct := UINT_TO_REAL(nTempU16) * 0.1;

(* ===== 协议输入 Byte 6-7: 实际焊接电流 (2字节小端, 0.1A分辨率) ===== *)
(* 范围: 0~400 对应0~400A *)
nTempU16 := BYTE_TO_UINT(GVL_Welders.g_byWeldIn[6]) + BYTE_TO_UINT(GVL_Welders.g_byWeldIn[7]) * 256;
GVL_Welders.g_rWeldCurrentAct := UINT_TO_REAL(nTempU16) * 0.1;

(* ===== 协议输入 Byte 8-9: 实际热丝焊接电流 (2字节小端, 10A分辨率) ===== *)
(* 范围: 0~20 对应0~200A *)
nTempU16 := BYTE_TO_UINT(GVL_Welders.g_byWeldIn[8]) + BYTE_TO_UINT(GVL_Welders.g_byWeldIn[9]) * 256;
GVL_Welders.g_rHotWireCurrentAct := UINT_TO_REAL(nTempU16) * 10.0;

(* ===== 协议输入 Byte 10-11: 送丝速度反馈 (已移除, 送丝通过轴控制) ===== *)

(* ===== 组装输入状态字 (PC通过D500读取) ===== *)
GVL_Welders.g_wWeldInStatus := 0;
IF GVL_Welders.g_bWeldArcOK      THEN GVL_Welders.g_wWeldInStatus := GVL_Welders.g_wWeldInStatus OR 16#0001; END_IF;
IF GVL_Welders.g_bWeldReady      THEN GVL_Welders.g_wWeldInStatus := GVL_Welders.g_wWeldInStatus OR 16#0002; END_IF;
IF GVL_Welders.g_bGunSwitchFault THEN GVL_Welders.g_wWeldInStatus := GVL_Welders.g_wWeldInStatus OR 16#0004; END_IF;
IF GVL_Welders.g_bWeldThermalProtect THEN GVL_Welders.g_wWeldInStatus := GVL_Welders.g_wWeldInStatus OR 16#0008; END_IF;
IF GVL_Welders.g_bWaterProtect   THEN GVL_Welders.g_wWeldInStatus := GVL_Welders.g_wWeldInStatus OR 16#0010; END_IF;
IF GVL_Welders.g_bWirePSThermal  THEN GVL_Welders.g_wWeldInStatus := GVL_Welders.g_wWeldInStatus OR 16#0020; END_IF;
IF GVL_Welders.g_bWirePSCommFault THEN GVL_Welders.g_wWeldInStatus := GVL_Welders.g_wWeldInStatus OR 16#0040; END_IF;
IF GVL_Welders.g_bWeldFault      THEN GVL_Welders.g_wWeldInStatus := GVL_Welders.g_wWeldInStatus OR 16#0080; END_IF;
IF GVL_Welders.g_bWeldHasCurrent     THEN GVL_Welders.g_wWeldInStatus := GVL_Welders.g_wWeldInStatus OR 16#0100; END_IF;

(* ================================================================ *)
(* D308 独立BOOL → 打包字 (PLC内部 → PC读D308)                         *)
(* CommPoll每周期从独立BOOL组装到g_wWeldStatusWord供PC读取             *)
(* ================================================================ *)
GVL_Welders.g_wWeldStatusWord := 0;
IF GVL_Welders.g_bWeldArcOK      THEN GVL_Welders.g_wWeldStatusWord := GVL_Welders.g_wWeldStatusWord OR 16#0001; END_IF;
IF GVL_Welders.g_bWeldReady      THEN GVL_Welders.g_wWeldStatusWord := GVL_Welders.g_wWeldStatusWord OR 16#0002; END_IF;
IF GVL_Welders.g_bWeldHasCurrent     THEN GVL_Welders.g_wWeldStatusWord := GVL_Welders.g_wWeldStatusWord OR 16#0004; END_IF;
IF GVL_Welders.g_bGunSwitchFault THEN GVL_Welders.g_wWeldStatusWord := GVL_Welders.g_wWeldStatusWord OR 16#0008; END_IF;
IF GVL_Welders.g_bWeldThermalProtect THEN GVL_Welders.g_wWeldStatusWord := GVL_Welders.g_wWeldStatusWord OR 16#0010; END_IF;
IF GVL_Welders.g_bWaterProtect   THEN GVL_Welders.g_wWeldStatusWord := GVL_Welders.g_wWeldStatusWord OR 16#0020; END_IF;
IF GVL_Welders.g_bWirePSThermal  THEN GVL_Welders.g_wWeldStatusWord := GVL_Welders.g_wWeldStatusWord OR 16#0040; END_IF;
IF GVL_Welders.g_bWirePSCommFault THEN GVL_Welders.g_wWeldStatusWord := GVL_Welders.g_wWeldStatusWord OR 16#0080; END_IF;
IF GVL_Welders.g_bWeldFault      THEN GVL_Welders.g_wWeldStatusWord := GVL_Welders.g_wWeldStatusWord OR 16#0100; END_IF;

END_PROGRAM
